(* PLC project Motor_Control, PLCAutoPilot Machine Expert Logic Builder V19.2.3.0, author PLCAutoPilot *)
(* stored: creationDateTime 2025-12-30T02:20:00.0000000, version 1.0.0.0, modificationDateTime 2025-12-30T02:20:00.0000000 *)

PROGRAM Motor_Control_LD
  VAR
    StartPB AT %IX0.0 : BOOL;
    StopPB AT %IX0.1 : BOOL;
    OverloadTrip AT %IX0.2 : BOOL;
    EmergencyStop AT %IX0.3 : BOOL;
    MotorContactor AT %QX0.0 : BOOL;
    RunIndicator AT %QX0.1 : BOOL;
    FaultIndicator AT %QX0.2 : BOOL;
  END_VAR
  VAR
    MotorRunning : BOOL;
    MotorFault : BOOL;
    SafetyOK : BOOL;
    StartCondition : BOOL;
    StartupTimer : TON;
  END_VAR

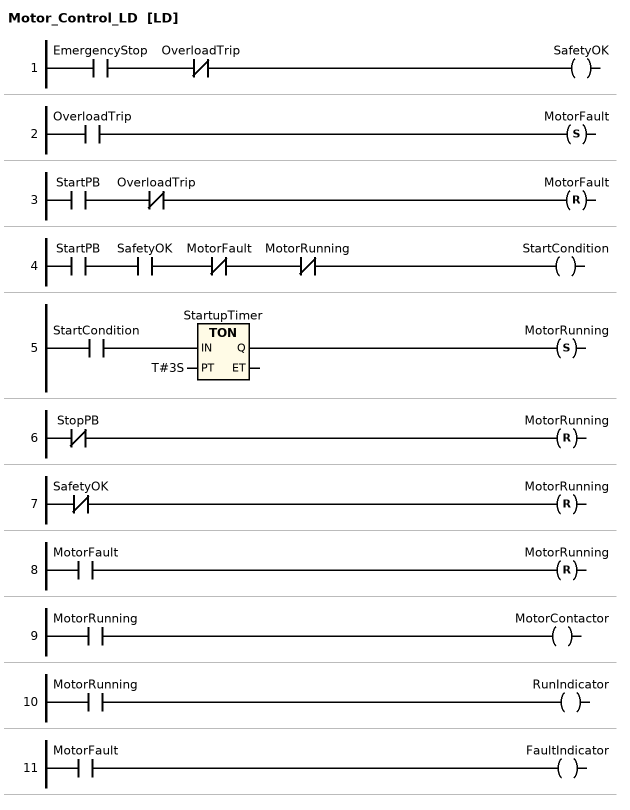
(* LD diagram, written out as Structured Text *)

SafetyOK := EmergencyStop AND NOT OverloadTrip;

IF OverloadTrip THEN MotorFault := TRUE; END_IF;

IF StartPB AND NOT OverloadTrip THEN MotorFault := FALSE; END_IF;

StartCondition := StartPB AND SafetyOK AND NOT MotorFault AND NOT MotorRunning;

StartupTimer(IN := StartCondition, PT := T#3S);
IF StartupTimer.Q THEN MotorRunning := TRUE; END_IF;

IF NOT StopPB THEN MotorRunning := FALSE; END_IF;

IF NOT SafetyOK THEN MotorRunning := FALSE; END_IF;

IF MotorFault THEN MotorRunning := FALSE; END_IF;

MotorContactor := MotorRunning;

RunIndicator := MotorRunning;

FaultIndicator := MotorFault;
END_PROGRAM
